(* PLC project case, CODESYS CODESYS V3.5 SP17 Patch 3 *)
(* stored: creationDateTime 2026-10-20T00:00:00 *)

PROGRAM PRG_A
  VAR
    xA : BOOL;
  END_VAR

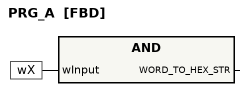
(* FBD diagram, written out as Structured Text *)
AND(wX);
END_PROGRAM

CONFIGURATION Device
  RESOURCE Application ON PLC
  END_RESOURCE
END_CONFIGURATION
